// TIA Portal V19 export
// export: Created 2026-10-16T08:35:17.7165193Z, ExportSetting WithDefaults, DisplayName Totally Integrated Automation Portal, DisplayVersion V19, DisplayName TIA Portal Openness, DisplayVersion V19, DisplayName TIA Portal Version Control Interface, DisplayVersion V19, DisplayName STEP 7 Professional, DisplayVersion V19, DisplayName STEP 7 Safety, DisplayVersion V19, DisplayName WinCC Basic/Comfort/Advanced, DisplayVersion V19, DisplayName WinCC Unified, DisplayVersion V19
TagTable "ROLL_TP900_Tags"
  ROLL_Heartbeat : DInt  (PLC tag ROLL_HMI.Heartbeat, ROLL_PLC, 1 s)
  ROLL_Connected : Bool  (PLC tag ROLL_HMI.Connected, ROLL_PLC, 1 s)
  ROLL_ManualFunction : Int  (PLC tag ROLL_HMI.ManualFunction, ROLL_PLC, 1 s)
  ROLL_GroundHeld : Bool  (PLC tag ROLL_HMI.GroundHeld, ROLL_PLC, 1 s)
  ROLL_WorkHeld : Bool  (PLC tag ROLL_HMI.WorkHeld, ROLL_PLC, 1 s)
  ROLL_SelectedProgram : Int  (PLC tag ROLL_HMI.SelectedProgram, ROLL_PLC, 1 s)
  ROLL_RecipeCommand : Int  (PLC tag ROLL_HMI.RecipeCommand, ROLL_PLC, 1 s)
  ROLL_RecipeRequest : DInt  (PLC tag ROLL_HMI.RecipeRequest, ROLL_PLC, 1 s)
  ROLL_RecipeAck : DInt  (PLC tag ROLL_HMI.RecipeAck, ROLL_PLC, 1 s)
  ROLL_RecipeError : Int  (PLC tag ROLL_HMI.RecipeError, ROLL_PLC, 1 s)
  ROLL_CurrentProgram : Int  (PLC tag ROLL_HMI.CurrentProgram, ROLL_PLC, 1 s)
  ROLL_ParameterRequest : DInt  (PLC tag ROLL_HMI.ParameterRequest, ROLL_PLC, 1 s)
  ROLL_ParameterAck : DInt  (PLC tag ROLL_HMI.ParameterAck, ROLL_PLC, 1 s)
  ROLL_ParameterDb : Int  (PLC tag ROLL_HMI.ParameterDb, ROLL_PLC, 1 s)
  ROLL_ParameterIndex : Int  (PLC tag ROLL_HMI.ParameterIndex, ROLL_PLC, 1 s)
  ROLL_ParameterValue : DInt  (PLC tag ROLL_HMI.ParameterValue, ROLL_PLC, 1 s)
  ROLL_ParameterCurrentValue : DInt  (PLC tag ROLL_HMI.ParameterCurrentValue, ROLL_PLC, 1 s)
  ROLL_ParameterSlotPresent : Bool  (PLC tag ROLL_HMI.ParameterSlotPresent, ROLL_PLC, 1 s)
  ROLL_ParameterError : Int  (PLC tag ROLL_HMI.ParameterError, ROLL_PLC, 1 s)
  ROLL_Dwell1Seconds : Int  (PLC tag ROLL_HMI.Dwell1Seconds, ROLL_PLC, 1 s)
  ROLL_Drain1Seconds : Int  (PLC tag ROLL_HMI.Drain1Seconds, ROLL_PLC, 1 s)
  ROLL_Ultrasound1 : Bool  (PLC tag ROLL_HMI.Ultrasound1, ROLL_PLC, 1 s)
  ROLL_Dwell2Seconds : Int  (PLC tag ROLL_HMI.Dwell2Seconds, ROLL_PLC, 1 s)
  ROLL_Drain2Seconds : Int  (PLC tag ROLL_HMI.Drain2Seconds, ROLL_PLC, 1 s)
  ROLL_Dwell3Seconds : Int  (PLC tag ROLL_HMI.Dwell3Seconds, ROLL_PLC, 1 s)
  ROLL_Drain3Seconds : Int  (PLC tag ROLL_HMI.Drain3Seconds, ROLL_PLC, 1 s)
  ROLL_Dry4Seconds : Int  (PLC tag ROLL_HMI.Dry4Seconds, ROLL_PLC, 1 s)
  ROLL_BasketMotion : Int  (PLC tag ROLL_HMI.BasketMotion, ROLL_PLC, 1 s)
  ROLL_BathLift : Bool  (PLC tag ROLL_HMI.BathLift, ROLL_PLC, 1 s)
  ROLL_ProcessTimer1Units : Int  (PLC tag ROLL_HMI.ProcessTimer1Units, ROLL_PLC, 1 s)
  ROLL_ProcessTimer2Units : Int  (PLC tag ROLL_HMI.ProcessTimer2Units, ROLL_PLC, 1 s)
  ROLL_KeyF1 : Bool  (PLC tag ROLL_HMI.KeyF[1], ROLL_PLC, 1 s)
  ROLL_KeyF2 : Bool  (PLC tag ROLL_HMI.KeyF[2], ROLL_PLC, 1 s)
  ROLL_KeyF3 : Bool  (PLC tag ROLL_HMI.KeyF[3], ROLL_PLC, 1 s)
  ROLL_KeyF4 : Bool  (PLC tag ROLL_HMI.KeyF[4], ROLL_PLC, 1 s)
  ROLL_KeyF5 : Bool  (PLC tag ROLL_HMI.KeyF[5], ROLL_PLC, 1 s)
  ROLL_KeyF6 : Bool  (PLC tag ROLL_HMI.KeyF[6], ROLL_PLC, 1 s)
  ROLL_KeyF7 : Bool  (PLC tag ROLL_HMI.KeyF[7], ROLL_PLC, 1 s)
  ROLL_KeyF8 : Bool  (PLC tag ROLL_HMI.KeyF[8], ROLL_PLC, 1 s)
  ROLL_KeyF9 : Bool  (PLC tag ROLL_HMI.KeyF[9], ROLL_PLC, 1 s)
  ROLL_KeyF10 : Bool  (PLC tag ROLL_HMI.KeyF[10], ROLL_PLC, 1 s)
  ROLL_KeyF11 : Bool  (PLC tag ROLL_HMI.KeyF[11], ROLL_PLC, 1 s)
  ROLL_KeyF12 : Bool  (PLC tag ROLL_HMI.KeyF[12], ROLL_PLC, 1 s)
  ROLL_KeyF13 : Bool  (PLC tag ROLL_HMI.KeyF[13], ROLL_PLC, 1 s)
  ROLL_KeyF14 : Bool  (PLC tag ROLL_HMI.KeyF[14], ROLL_PLC, 1 s)
  ROLL_KeyF15 : Bool  (PLC tag ROLL_HMI.KeyF[15], ROLL_PLC, 1 s)
  ROLL_KeyF16 : Bool  (PLC tag ROLL_HMI.KeyF[16], ROLL_PLC, 1 s)
  ROLL_Clock : Bool  (PLC tag ROLL_HMI.StatusM[3,5], ROLL_PLC, 100 ms)
  ROLL_ManualMode : Bool  (PLC tag ROLL_IO.Input[0,1], ROLL_PLC, 1 s)
  ROLL_Simulation : Bool  (PLC tag ROLL_IO.Simulation, ROLL_PLC, 1 s)
  ROLL_OutputsEnabled : Bool  (PLC tag ROLL_IO.PhysicalOutputsEnabled, ROLL_PLC, 1 s)
  ROLL_IoConfigured : Bool  (PLC tag ROLL_IO.PhysicalIoConfigured, ROLL_PLC, 1 s)
  ROLL_ConversionFault : Bool  (PLC tag ROLL_IO.ConversionFault, ROLL_PLC, 1 s)
